(* IEC 61131-3 sources: nautilus/internal/project/testdata/libdir/hmi, 1 file *)

(* ---- ignored.st ---- *)
FUNCTION_BLOCK HiAlarm
VAR_INPUT PV : REAL; END_VAR
END_FUNCTION_BLOCK
